(* IEC 61131-3 sources: IRIS-Project/LASAL CONTROL SOFTWARE/LasalProject_2025_09_12/Class/DischargeTimer, 1 file *)

(* ---- DischargeTimer.st ---- *)
(*!
<Class
	Name               = "DischargeTimer"
	Revision           = "0.0"
	RealtimeTask       = "false"
	CyclicTask         = "true"
	DefCyclictime      = "100 ms"
	BackgroundTask     = "false"
	Sigmatek           = "false"
	OSInterface        = "false"
	HighPriority       = "false"
	Automatic          = "false"
	UpdateMode         = "Prescan"
	SharedCommandTable = "true"
	Objectsize         = "(530,120)">
	<Channels>
		<Server Name="ClassSvr" Visualized="false" Initialize="false" WriteProtected="true" Retentive="false"/>
		<Server Name="s_DisTimer1" Visualized="false" Initialize="false" WriteProtected="false" Retentive="false"/>
		<Server Name="s_DisTimer2" Visualized="false" Initialize="false" WriteProtected="false" Retentive="false"/>
		<Server Name="s_DisTimer3" Visualized="false" Initialize="false" WriteProtected="false" Retentive="false"/>
		<Server Name="s_Reset" Visualized="false" Initialize="false" WriteProtected="false" Retentive="false"/>
		<Server Name="s_StartStopTimer" Visualized="false" Initialize="false" WriteProtected="false" Retentive="false"/>
		<Client Name="c_SysDate" Required="true" Internal="false"/>
		<Client Name="c_SysTime" Required="true" Internal="false"/>
		<Client Name="c_timer" Required="true" Internal="false"/>
	</Channels>
</Class>
*)
DischargeTimer : CLASS
  //Servers:
	ClassSvr 	: SvrChCmd_DINT;
	s_StartStopTimer 	: SvrCh_DINT;
	s_DisTimer1 	: SvrCh_DINT;
	s_DisTimer2 	: SvrCh_DINT;
	s_DisTimer3 	: SvrCh_DINT;
	s_Reset 	: SvrCh_DINT;
  //Clients:
	c_timer 	: CltChCmd_TimeDateLib;
	c_SysDate 	: CltCh_DINT;
	c_SysTime 	: CltCh_TIME_LSL;
  //Variables:
		v_hd_Date 	: HDINT;
		v_hd_Time_1 	: HDINT;
		v_day 	: UDINT;
		v_month 	: UDINT;
		v_year 	: UDINT;
		v_hd_Time_2 	: HDINT;
		case_Time 	: DINT;
		v_tot_seconds 	: DINT;
		v_tot_minutes 	: DINT;
		a 	: DINT;
		i 	: DINT;
  //Functions:

	FUNCTION VIRTUAL GLOBAL Init;

	FUNCTION VIRTUAL GLOBAL CyWork
		VAR_INPUT
			EAX 	: UDINT;
		END_VAR
		VAR_OUTPUT
			state (EAX) 	: UDINT;
		END_VAR;
  //Tables:
	FUNCTION @STD
		VAR_OUTPUT
			ret_code	: CONFSTATES;
		END_VAR;
	FUNCTION GLOBAL TAB @CT_;
END_CLASS;

#pragma usingLtd TimeDateLib

FUNCTION VIRTUAL GLOBAL DischargeTimer::CyWork
	VAR_INPUT
		EAX 	: UDINT;
	END_VAR
	VAR_OUTPUT
		state (EAX) 	: UDINT;
	END_VAR

  //READ ACTUAL TIME AND DATE FROM CLIENTS; shr for shift bits
  //v_hd_Date := c_SysDate.Read();
  //v_hd_Time_1 := c_SysTime.Read();

  ///v_seconds_1 := (v_hd_Time_1 AND 16#0000FF00) shr 8;
  //v_minutes_1 := (v_hd_Time_1 AND 16#00FF0000) shr 16;
  //v_hours_1   := (v_hd_Time_1 AND 16#FF000000) shr 24;

  //v_day     := (v_hd_Date AND 16#00000FF0) shr 4;
  //v_month   := (v_hd_Date AND 16#0000F000) shr 12;
  //v_year    := (v_hd_Date AND 16#FFFF0000) shr 16;

  if s_Reset.Read() then
     s_DisTimer1.Write(input:=0);
     s_DisTimer2.Write(input:=0);
     s_DisTimer3.Write(input:=0);
     i:=0;
     case_Time:=0;
  end_if;

  case case_Time of

    0:
      if s_StartStopTimer.Read() then
        v_hd_Time_1 := c_SysTime.Read();
        case_Time:=10;
      end_if;

    10:
      if s_StartStopTimer.Read()=0 then
        v_hd_Time_2 := c_SysTime.Read();
        case_Time:=20;
      end_if;

    20:
      v_tot_seconds := c_timer.TimeDiff(tim1:=v_hd_Time_2, tim2:=v_hd_Time_1);
      case_Time:=30;

    30:

      v_tot_minutes :=v_tot_seconds / 60; //minuti
      a := v_tot_seconds mod 60; //secondi
      i+=1;
      case_Time:=40;

     40:

      case i of
        0:

        1:
          s_DisTimer1.Write(input:=v_tot_seconds);
          case_Time:=0;
        2:
          s_DisTimer2.Write(input:=v_tot_seconds);
          case_Time:=0;
        3:
          s_DisTimer3.Write(input:=v_tot_seconds);
          case_Time:=50;

      end_case;

    50:

  end_case;

	state := READY;

END_FUNCTION

FUNCTION VIRTUAL GLOBAL DischargeTimer::Init

END_FUNCTION
